// TIA Portal V19 export
TYPE "ST_DOOR"
   STRUCT
      SafetyDoors_Locked : Bool;
      SafetyDoor_1 : Bool;
      SafetyDoor_2 : Bool;
      SafetyDoor_3 : Bool;
      SafetyDoor_4 : Bool;
      SafetyDoor_5 : Bool;
      SafetyDoor_6 : Bool;
      SafetyDoor_7 : Bool;
      SafetyDoor_8 : Bool;
      SafetyDoor_9 : Bool;
      SafetyDoor_10 : Bool;
   END_STRUCT;
END_TYPE
